FUNCTION_BLOCK SimulationCheck IMPLEMENTS I_Diagnosable
VAR
    _IsOnMachine    : BOOL;
    _NotFinalCount  : DINT;
    _NotFinalNames  : STRING(255);
END_VAR
(*
    SimulationCheck

    Told, while wiring, the name and source of every routed device. Lists
    every device that isn't FinalHardware, for the HMI and the event log.
    On a controller whose site is the machine itself, each of them is a
    fault.
*)

METHOD FB_init : BOOL
VAR_INPUT
    bInitRetains : BOOL;
    bInCopyCode  : BOOL;
    IsOnMachine  : BOOL;
END_VAR
_IsOnMachine := IsOnMachine;
END_METHOD

METHOD PUBLIC AddDevice : BOOL
VAR_INPUT
    Name   : STRING(32);
    Source : E_DeviceSource;
END_VAR
AddDevice := TRUE;
IF Source = E_DeviceSource.FinalHardware THEN
    RETURN;
END_IF
_NotFinalCount := _NotFinalCount + 1;
IF _NotFinalCount = 1 THEN
    _NotFinalNames := Name;
ELSE
    _NotFinalNames := CONCAT(CONCAT(_NotFinalNames, ', '), Name);
END_IF
END_METHOD

PROPERTY PUBLIC Name : STRING
GET
Name := 'Device sources';
END_GET
END_PROPERTY

PROPERTY PUBLIC HasFault : BOOL
GET
HasFault := _IsOnMachine AND _NotFinalCount > 0;
END_GET
END_PROPERTY

PROPERTY PUBLIC FaultText : STRING
GET
IF HasFault THEN
    FaultText := CONCAT('Not final hardware: ', _NotFinalNames);
ELSE
    FaultText := '';
END_IF
END_GET
END_PROPERTY

PROPERTY PUBLIC NotFinalDevices : STRING(255)
GET
NotFinalDevices := _NotFinalNames;
END_GET
END_PROPERTY

PROPERTY PUBLIC NotFinalCount : DINT
GET
NotFinalCount := _NotFinalCount;
END_GET
END_PROPERTY

END_FUNCTION_BLOCK

(* stored: Version 1.1.0.1, ProductVersion 3.1.4026.0
   POU SimulationCheck: Id {f75636c3-6bcd-4d43-a3d8-a0d96221c0ba}, SpecialFunc None
   Folder I_Diagnosable: Id {78fc4a9a-42f6-4515-8c65-c7673cf49001}
   Method FB_init: Id {fea14d57-7242-403b-80fd-74771c8419eb}
   Method AddDevice: Id {b3c2d89d-1d54-4319-af9c-0b55c47b7405}
   Property Name: Id {2801ce61-39a9-4109-8621-2fc2fa85c6b6}
   Get Get: Id {e7e29e38-246f-4901-bc44-042893e44680}
   Property HasFault: Id {158cb11b-d26a-479c-8bc2-bebef980beb6}
   Get Get: Id {428a8075-6a87-40ea-b295-78a1cea1da50}
   Property FaultText: Id {b53d9a1b-9674-444f-92e0-382c5b28911b}
   Get Get: Id {ff55fe03-c039-462d-bb89-10b82e575e47}
   Property NotFinalDevices: Id {70d9c4e2-997d-4b99-9043-8feae373cf66}
   Get Get: Id {8cfc2eca-0657-487b-8b80-4af77d2befe5}
   Property NotFinalCount: Id {d154facf-767b-4c4b-96d3-b0f059226c59}
   Get Get: Id {5f6d15aa-c349-4627-809b-ffe0d6dd37d5} *)
